// TIA Portal V20 export
Screen "160PRBCompleteDisplay_1"  1276x673
  ScreenItem "Title_ScreenOverview_X390_Y2" at 390,2 size 500x30  Type=HmiTextBox
  ScreenItem "Button_Back_1" at 2,2 size 90x60  Type=HmiButton
  ScreenItem "sequenceControlFaceplate_Lite_1" at 383,557 size 641x64  Type=HmiFaceplateContainer
  ScreenItem "Line_Header_X0_Y64" at 0,64 size 1276x0  Type=HmiLine
  ScreenItem "permanentareaborderrectangle" at 0,0 size 0x0  Type=HmiRectangle
  ScreenItem "Button_Back" at 2,4 size 90x60  Type=HmiButton
  ScreenItem "Title_ScreenOverview_X390_Y2_1" at 380,5 size 510x57  Type=HmiTextBox
  ScreenItem "Button_Back_2" at 1171,612 size 90x60  Type=HmiButton
  ScreenItem "Move_Legend" at 1182,2 size 90x60  Type=HmiButton
  ScreenItem "面板容器_1" at 12,276 size 163x70  Type=HmiFaceplateContainer
  ScreenItem "面板容器_4" at 12,344 size 163x70  Type=HmiFaceplateContainer
  ScreenItem "面板容器_3" at 195,276 size 163x70  Type=HmiFaceplateContainer
  ScreenItem "面板容器_11" at 436,276 size 163x70  Type=HmiFaceplateContainer
  ScreenItem "面板容器_12" at 857,276 size 163x70  Type=HmiFaceplateContainer
  ScreenItem "面板容器_2" at 1090,4 size 88x58  Type=HmiFaceplateContainer
  ScreenItem "OPMode4_Foreground_Blocked" at 1090,4 size 88x58  Type=HmiGraphicView
